{attribute 'Tc2GvlVarNames'}
VAR_GLOBAL
	stgGr05Alarm			:ST_AlarmRef;
END_VAR

(* stored: Version 1.1.0.1, ProductVersion 3.1.4024.15
   GVL GVL_Gr05Alarm: Id {8ab8aab8-2f53-4d48-b697-72ac4fd77c00} *)
